Fanuc KAREL source: ko00090.KL

-- PROVISIONAL review KL for V1013-1; original PC SHA256 e0f59b9ff963bb4234059738d214da79cc3039b1bcf45f8cd4f8e18074b8efb7
-- Incomplete behavior may be omitted. Consult companion uncertainty JSON. Do not deploy.
PROGRAM KO00090
%NOLOCKGROUP
BEGIN
  -- UNRESOLVED_PC offsets 5-12; opcodes 9D,23
  -- UNRESOLVED_PC offsets 17-69; opcodes 27,27,49,7E,AD,27,49,7E,AD,22,31,7E,4A
  -- UNRESOLVED_PC offsets 74-78; opcodes 7F
END KO00090
